// TIA Portal V20 export
// export: Created 2026-10-11T05:28:41.5387806Z, ExportSetting WithDefaults, DisplayName Totally Integrated Automation Portal, DisplayVersion V20, DisplayName TIA Portal Openness, DisplayVersion V20, DisplayName TIA Portal Teamcenter Gateway, DisplayVersion V20, DisplayName TIA Portal Version Control Interface, DisplayVersion V20, DisplayName SINAMICS Startdrive Advanced, DisplayVersion V20 SP1 Update 2, DisplayName SINAMICS Startdrive G110M, G120, G120C, G120D, G120P, G115D, DisplayVersion V20 SP1 Update 2, DisplayName SINAMICS Startdrive G130, G150, S120, S150, SINAMICS MV, G220, S200, S210, DisplayVersion V20 SP1 Update 2, DisplayName STEP 7 Professional, DisplayVersion V20, DisplayName STEP 7 Safety, DisplayVersion V20, DisplayName WinCC Basic/Comfort/Advanced, DisplayVersion V20, DisplayName WinCC Professional, DisplayVersion V20, DisplayName WinCC Unified, DisplayVersion V20
TYPE "ST_HmiResponse"
// stored: IsFailsafeCompliant false
   STRUCT
      AckSequence : UDInt;
      Accepted : Bool;
      Diagnostic : WString[255];
      Report { S7_SetPoint := 'True'} : "ST_ReleaseReport";
      ConfigPage { S7_SetPoint := 'True'} : "ST_ConfigPage";
   END_STRUCT;
END_TYPE
